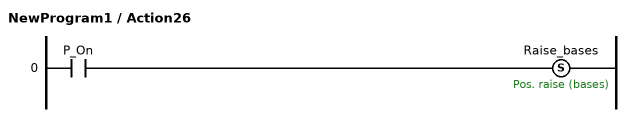
; [picture p24: NewProgram1 / Action26, rungs 0-0]
; rung 0
LD P_On
SET Raise_bases  ; Pos. raise (bases)

### Action Action27

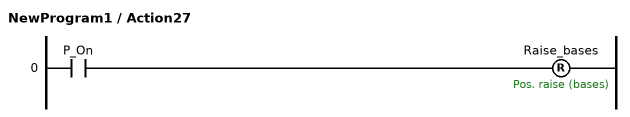
; rung 0
LD P_On
RSET Raise_bases  ; Pos. raise (bases)

### Action Action28

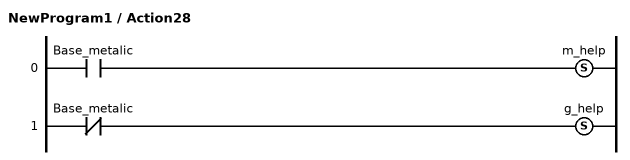
; rung 0
LD Base_metalic
SET m_help
; rung 1
LDNOT Base_metalic
SET g_help

## Program NewProgram2 (cyclic task 1)
IF P_First_Cycle THEN
	g_num := 11;
	m_num := 12;
	(*g_comp := FALSE;*)
	m_comp := FALSE;
	g_help:= FALSE;
	m_help:= FALSE;
	
	g_comp := TRUE;
END_IF;





IF (g_num / 10) = 0 THEN
	g_comp:=TRUE;
END_IF;

IF g_comp AND m_comp THEN
	Stop_light := True;
	
END_IF;

IF (m_num / 10) = 0 THEN
	m_comp:=TRUE;
	g_comp:= FALSE;
END_IF;

IF m_help THEN
	m_num:= m_num - 10;
	m_help:= FALSE;
ELSIF g_help THEN
	g_num:= g_num - 10;
	g_help:= FALSE;
END_IF;
	

## Program NewProgram3 (cyclic task 2)
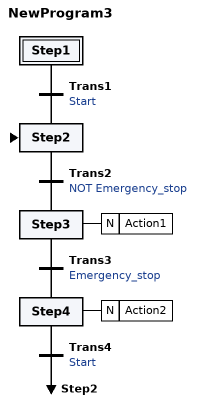
INITIAL_STEP Step1 :
END_STEP
TRANSITION Trans1 FROM Step1 TO Step2
 := Start;
END_TRANSITION
STEP Step2 :
END_STEP
TRANSITION Trans2 FROM Step2 TO Step3
 := NOT Emergency_stop;
END_TRANSITION
STEP Step3 :
Action1(N) ;
END_STEP
TRANSITION Trans3 FROM Step3 TO Step4
 := Emergency_stop;
END_TRANSITION
STEP Step4 :
Action2(N) ;
END_STEP
TRANSITION Trans4 FROM Step4 TO Step2
 := Start;
END_TRANSITION

### Action Action1

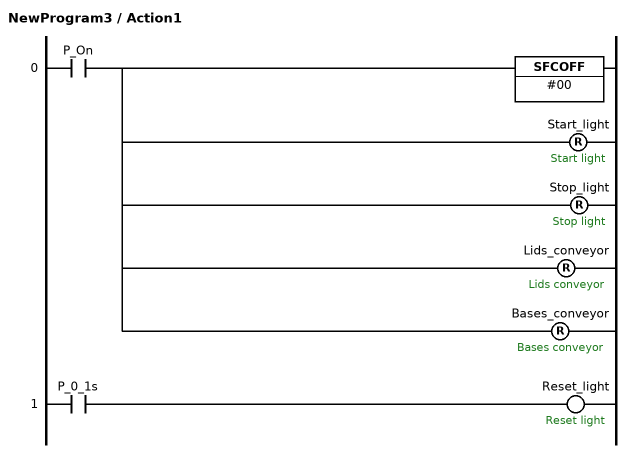
; rung 0
LD P_On
SFCOFF #00
RSET Start_light  ; Start light
RSET Stop_light  ; Stop light
RSET Lids_conveyor  ; Lids conveyor
RSET Bases_conveyor  ; Bases conveyor
; rung 1
LD P_0_1s
OUT Reset_light  ; Reset light

### Action Action2

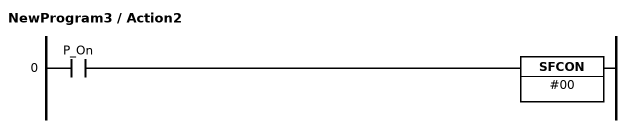
; rung 0
LD P_On
SFCON #00